Fanuc KAREL source: KB00130.KL

PROGRAM KB00130
%NOLOCKGROUP
%ENVIRONMENT MULTI
VAR
  P1: INTEGER
  P2: INTEGER
  P3: BOOLEAN
BEGIN
  P1 = 1
  P2 = 1
  P3 = TRUE
  PEND_SEMA(P1, P2, P3)
END KB00130
